// TwinCAT 3 PLC project PLCStudent
// ProgramVersion: 3.1.4026.20
// libraries:
//   Tc2_Standard, * (Beckhoff Automation GmbH)
//   Tc2_System, * (Beckhoff Automation GmbH)
//   Tc3_Module, * (Beckhoff Automation GmbH)
// project tree:
//   GVLs/ GVL.TcGVL
//   / PlcTask.TcTTO
//   POUs/ Control_FBD.TcPOU, MAIN.TcPOU
// (motion and I/O tree: see PLC project plcsim)
// real-time tasks:
//   TASK PlcTask: cycle T#20ms, priority 20, ADS port 350
// variable links:
//   PLCSim/PLCSim Instance <-> PLCStudent/PLCStudent Instance
//     PlcTask Inputs/GVL.ixDoorClose <-> PlcTask Outputs/GVL.qxDoorClose
//     PlcTask Inputs/GVL.ixLampElevat1 <-> PlcTask Outputs/GVL.qxLampElevat1
//     PlcTask Inputs/GVL.ixLampElevat2 <-> PlcTask Outputs/GVL.qxLampElevat2
//     PlcTask Inputs/GVL.ixLampElevat3 <-> PlcTask Outputs/GVL.qxLampElevat3
//     PlcTask Inputs/GVL.ixLampLevel1 <-> PlcTask Outputs/GVL.qxLampLevel1
//     PlcTask Inputs/GVL.ixLampLevel2 <-> PlcTask Outputs/GVL.qxLampLevel2
//     PlcTask Inputs/GVL.ixLampLevel3 <-> PlcTask Outputs/GVL.qxLampLevel3
//     PlcTask Inputs/GVL.ixMotorDown <-> PlcTask Outputs/GVL.qxMotorDown
//     PlcTask Inputs/GVL.ixMotorUp <-> PlcTask Outputs/GVL.qxMotorUp
//     PlcTask Outputs/GVL.qxButtElevat1 <-> PlcTask Inputs/GVL.ixButtElevat1
//     PlcTask Outputs/GVL.qxButtElevat2 <-> PlcTask Inputs/GVL.ixButtElevat2
//     PlcTask Outputs/GVL.qxButtElevat3 <-> PlcTask Inputs/GVL.ixButtElevat3
//     PlcTask Outputs/GVL.qxButtGreen <-> PlcTask Inputs/GVL.ixButtGreen
//     PlcTask Outputs/GVL.qxButtLevel1 <-> PlcTask Inputs/GVL.ixButtLevel1
//     PlcTask Outputs/GVL.qxButtLevel2 <-> PlcTask Inputs/GVL.ixButtLevel2
//     PlcTask Outputs/GVL.qxButtLevel3 <-> PlcTask Inputs/GVL.ixButtLevel3
//     PlcTask Outputs/GVL.qxButtRed <-> PlcTask Inputs/GVL.ixButtRed
//     PlcTask Outputs/GVL.qxDoorClosed <-> PlcTask Inputs/GVL.ixDoorClosed
//     PlcTask Outputs/GVL.qxDoorOpen <-> PlcTask Inputs/GVL.ixDoorOpen
//     PlcTask Outputs/GVL.qxElevatLevel1 <-> PlcTask Inputs/GVL.ixElevatLevel1
//     PlcTask Outputs/GVL.qxElevatLevel2 <-> PlcTask Inputs/GVL.ixElevatLevel2
//     PlcTask Outputs/GVL.qxElevatLevel3 <-> PlcTask Inputs/GVL.ixElevatLevel3

CONFIGURATION PLCStudent
    RESOURCE PLC ON TwinCAT3
        TASK PlcTask(INTERVAL := T#20ms, PRIORITY := 20);
        PROGRAM MAIN WITH PlcTask : MAIN;
    END_RESOURCE
END_CONFIGURATION

// ---- GVLs/GVL.TcGVL
{attribute 'qualified_only'}
VAR_GLOBAL
//Input to PLC from process
	ixButtLevel1		AT %I*:	BOOL;		(* Button at level 1 *)
	ixButtLevel2		AT %I*:	BOOL;		(* Button at level 2 *)
	ixButtLevel3		AT %I*:	BOOL;		(* Button at level 3 *)

	ixElevatLevel1 		AT %I*: BOOL;		(* Sensor at level 1 for elevator presence *)
	ixElevatLevel2 		AT %I*: BOOL;		(* Sensor at level 2 for elevator presence *)
	ixElevatLevel3 		AT %I*: BOOL;		(* Sensor at level 3 for elevator presence *)

	ixButtGreen 		AT %I*:	BOOL;		(* Green button *)
	ixButtRed			AT %I*:	BOOL;		(* Red button, normally closed *)

	ixButtElevat1		AT %I*:	BOOL;		(* Button 1 inside elevator PLCSim only *)
	ixButtElevat2		AT %I*:	BOOL;		(* Button 2 inside elevator PLCSim only *)
	ixButtElevat3		AT %I*:	BOOL;		(* Button 3 inside elevator PLCSim only *)
	
	ixDoorClosed		AT %I*: BOOL;		(* Sensor for door closed PLCSim only *)
	ixDoorOpen			AT %I*:	BOOL;		(* Sensor for door open   PLCSim only *)

//Output from PLC to process
	qxLampLevel1		AT %Q*:	BOOL;		(* Lamp at level 1*)
	qxLampLevel2		AT %Q*:	BOOL;		(* Lamp at level 2*)
	qxLampLevel3		AT %Q*:	BOOL;		(* Lamp at level 3*)
	qxMotorDown			AT %Q*:	BOOL;		(* Run motor down *)
	qxMotorUp			AT %Q*:	BOOL;		(* Run motor up *)

	qxLampElevat1 		AT %Q*:	BOOL;		(* Lamp 1 inside elevator PLCSim only*)
	qxLampElevat2 		AT %Q*:	BOOL;		(* Lamp 2 inside elevator PLCSim only *)
	qxLampElevat3 		AT %Q*:	BOOL;		(* Lamp 3 inside elevator PLCSim only *)

	qxDoorClose			AT %Q*:	BOOL;		(* Close door and keep it closed  PLCSim only *)
	qiDispElevat 		AT %Q*:	UINT;		(* Integer display inside elevator PLCSim only *)
END_VAR

// ---- POUs/MAIN.TcPOU
PROGRAM MAIN
VAR
END_VAR

Control_FBD();

END_PROGRAM

// ---- POUs/Control_FBD.TcPOU
PROGRAM Control_FBD
VAR
	
	batLevel1 : BOOL;
	batLevel2: BOOL;
	batLevel3: BOOL;
	
	mxRun : BOOL;
	qxMotorUp : BOOL;
	qxMotorDown: BOOL;
	
	SR1: SR;
	RS1: RS;
	TOF_1: TOF;
	TON_1: TON;
END_VAR
VAR // added by the converter: edge detectors and wires of the graphical bodies
    _w1, _w2, _w3 : BOOL;
END_VAR

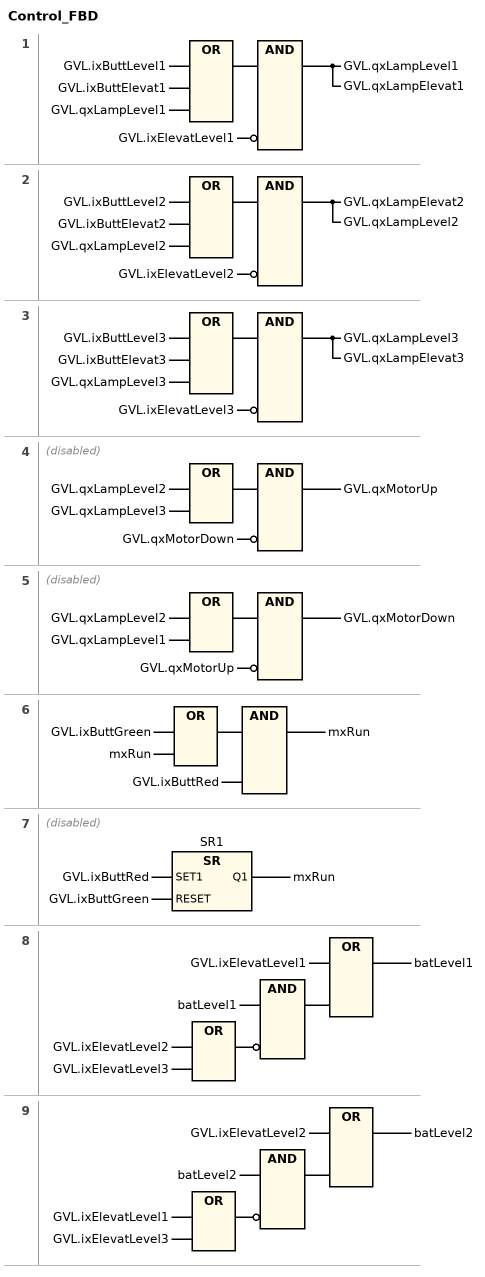
// NETWORK 1
_w1 := (GVL.ixButtLevel1 OR GVL.ixButtElevat1 OR GVL.qxLampLevel1) AND NOT GVL.ixElevatLevel1;
GVL.qxLampLevel1 := _w1;
GVL.qxLampElevat1 := _w1;

// NETWORK 2
_w2 := (GVL.ixButtLevel2 OR GVL.ixButtElevat2 OR GVL.qxLampLevel2) AND NOT GVL.ixElevatLevel2;
GVL.qxLampElevat2 := _w2;
GVL.qxLampLevel2 := _w2;

// NETWORK 3
_w3 := (GVL.ixButtLevel3 OR GVL.ixButtElevat3 OR GVL.qxLampLevel3) AND NOT GVL.ixElevatLevel3;
GVL.qxLampLevel3 := _w3;
GVL.qxLampElevat3 := _w3;

// NETWORK 4 (disabled)
// GVL.qxMotorUp := (GVL.qxLampLevel2 OR GVL.qxLampLevel3) AND NOT GVL.qxMotorDown;

// NETWORK 5 (disabled)
// GVL.qxMotorDown := (GVL.qxLampLevel2 OR GVL.qxLampLevel1) AND NOT GVL.qxMotorUp;

// NETWORK 6
mxRun := (GVL.ixButtGreen OR mxRun) AND GVL.ixButtRed;

// NETWORK 7 (disabled)
// SR1(SET1 := GVL.ixButtRed, RESET := GVL.ixButtGreen); // SR
// mxRun := SR1.Q1;

// NETWORK 8
batLevel1 := GVL.ixElevatLevel1 OR batLevel1 AND NOT (GVL.ixElevatLevel2 OR GVL.ixElevatLevel3);

// NETWORK 9
batLevel2 := GVL.ixElevatLevel2 OR batLevel2 AND NOT (GVL.ixElevatLevel1 OR GVL.ixElevatLevel3);

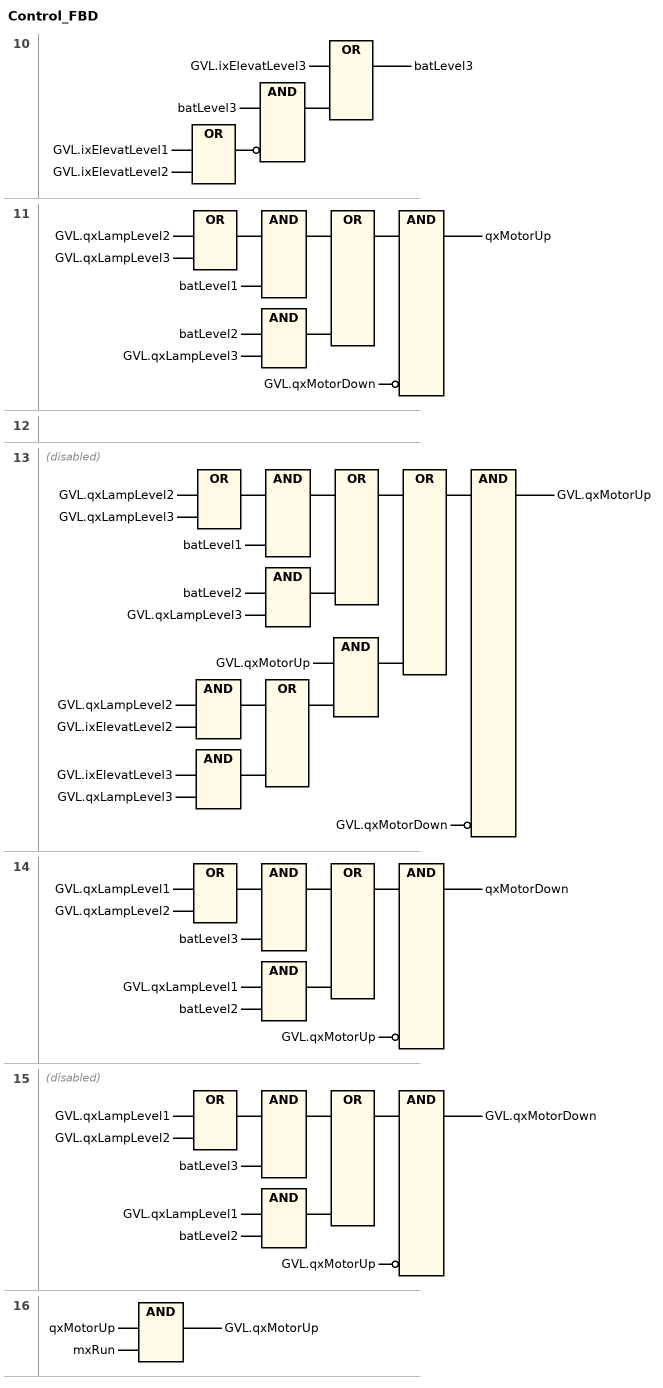
// NETWORK 10
batLevel3 := GVL.ixElevatLevel3 OR batLevel3 AND NOT (GVL.ixElevatLevel1 OR GVL.ixElevatLevel2);

// NETWORK 11
qxMotorUp := ((GVL.qxLampLevel2 OR GVL.qxLampLevel3) AND batLevel1 OR batLevel2 AND GVL.qxLampLevel3) AND NOT GVL.qxMotorDown;

// NETWORK 12

// NETWORK 13 (disabled)
// GVL.qxMotorUp := (((GVL.qxLampLevel2 OR GVL.qxLampLevel3) AND batLevel1 OR batLevel2 AND GVL.qxLampLevel3) OR GVL.qxMotorUp AND (GVL.qxLampLevel2 AND GVL.ixElevatLevel2 OR GVL.ixElevatLevel3 AND GVL.qxLampLevel3)) AND NOT GVL.qxMotorDown;

// NETWORK 14
qxMotorDown := ((GVL.qxLampLevel1 OR GVL.qxLampLevel2) AND batLevel3 OR GVL.qxLampLevel1 AND batLevel2) AND NOT GVL.qxMotorUp;

// NETWORK 15 (disabled)
// GVL.qxMotorDown := ((GVL.qxLampLevel1 OR GVL.qxLampLevel2) AND batLevel3 OR GVL.qxLampLevel1 AND batLevel2) AND NOT GVL.qxMotorUp;

// NETWORK 16
GVL.qxMotorUp := qxMotorUp AND mxRun;

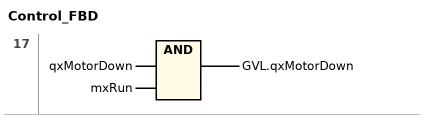
// NETWORK 17
GVL.qxMotorDown := qxMotorDown AND mxRun;

END_PROGRAM
